Fanuc KAREL source: kt00549.KL

-- PROVISIONAL review KL for V940-1; original PC SHA256 e77ba5bfc8690790f66ef0cc53d7b1d036eafe68abb5a4e96473a725d4199116
-- Incomplete behavior may be omitted. Consult companion uncertainty JSON. Do not deploy.
PROGRAM KT00549
%NOLOCKGROUP
-- UNRESOLVED_DECL P1 type=000199
-- UNRESOLVED_DECL P2 type=000199
-- UNRESOLVED_DECL OUT type=000101
BEGIN
  -- V9_ZERO_TABLE_METADATA_HINT layout=0001; no indexed target words; source/name/runtime held
  -- UNRESOLVED_PC offsets 5-39; opcodes 49,7E,49,7E,60,4A
  -- UNRESOLVED_PC offsets 44-48; opcodes 7F
END KT00549
